(* Logix 5000 project; controller SmartManufacturingCell Emulate 5570 rev 33.11; software revision 33.03 *)
// Simulation only. Core cell candidate; acceptance pending.

TASK MainTask (periodic, rate 20 ms, priority 10, watchdog 500 ms) : Program_System, Program_Conveyor, Program_Filling, Program_Inspection, Program_Production, Program_Simulation

MODULES
   Local : Emulate 5570 (ICP 4, rev 33.11)
END_MODULES

TYPE UDT_Bottle :   // Bottle record
STRUCT
   Occupied : BOOL;   // A tracked bottle occupies this position
   FillComplete : BOOL;   // This bottle completed filling
   InspectionComplete : BOOL;   // This bottle has a valid inspection result
   RejectRequired : BOOL;   // Inspection determined this bottle must be rejected
END_STRUCT
END_TYPE

VAR_GLOBAL   (* controller tags *)
   Cfg_FillTimeMs : DINT := 1500;   // Fill duration; 100..3000 ms. Sampled when filling starts.
   Cfg_InspectionTimeMs : DINT := 500;   // Inspection duration; 100..2000 ms. Sampled when inspection starts.
   Conveyor_Flt_FailToStart : BOOL; {access Read Only}   // Conveyor commanded but running feedback missing for 2 s Latched; clear cell, remove cause, then fresh Reset.
   Conveyor_Sts_ResetAccepted : BOOL; {access Read Only}   // One-execution indication that conveyor fault reset was accepted.
   Exit_Flt_DischargeTimeout : BOOL; {access Read Only}   // Good or reject bottle departure not confirmed within 3 s Latched; clear cell, remove cause, then fresh Reset.
   Exit_Sts_GoodCompletePulse : BOOL; {access Read Only}   // Exit Sts GoodCompletePulse
   Exit_Sts_RejectCompletePulse : BOOL; {access Read Only}   // Exit Sts RejectCompletePulse
   Exit_Sts_ResetAccepted : BOOL; {access Read Only}   // Exit Sts ResetAccepted
   Exit_Sts_State : DINT; {access Read Only}   // 0 Empty; 10 Waiting; 20 Good discharge; 30 Extending; 40 Reject discharge; 50 Retracting; 60 Complete; 90 Faulted
   Filling_Flt_FillTimeout : BOOL; {access Read Only}   // Fill completion not received within 4 s Latched; clear cell, remove cause, then fresh Reset.
   Filling_Flt_ValveFailToClose : BOOL; {access Read Only}   // Fill valve did not close within 2 s Latched; clear cell, remove cause, then fresh Reset.
   Filling_Sts_ActiveFillTimeMs : DINT; {access Read Only}   // Sampled fill duration for current bottle
   Filling_Sts_ResetAccepted : BOOL; {access Read Only}   // Filling Sts ResetAccepted
   Filling_Sts_State : DINT; {access Read Only}   // 0 Empty; 10 Waiting; 20 Filling; 30 Closing; 40 Complete; 90 Faulted
   HMI_Cmd_Acknowledge : BOOL;   // Acknowledge alarm indication; does not reset faults
   HMI_Cmd_ClearCell : BOOL;   // Request removal of simulated bottles during fault recovery
   HMI_Cmd_ConveyorJog : BOOL;   // Request conveyor movement while held
   HMI_Cmd_FillValveOpen : BOOL;
   HMI_Cmd_LoadBottle : BOOL;   // Request one simulated bottle at the available entry position
   HMI_Cmd_RejectExtend : BOOL;
   HMI_Cmd_Reset : BOOL;   // Request fault reset after recovery conditions are satisfied
   HMI_Cmd_ResetStatistics : BOOL;   // Clear production statistics only when Stopped and cell empty
   HMI_Cmd_SelectAuto : BOOL;   // Request Auto mode
   HMI_Cmd_SelectManual : BOOL;   // Request Manual mode
   HMI_Cmd_Start : BOOL;   // Request automatic production start
   HMI_Cmd_Stop : BOOL;   // Request controlled production stop
   HMI_Sim_BottleMissingAtFill : BOOL;   // Suppress Fill photoeye while retaining simulated bottle presence. Simulation test only.
   HMI_Sim_ConveyorFailToStart : BOOL;   // Suppress conveyor running feedback. Simulation test only.
   HMI_Sim_FillFailToComplete : BOOL;   // Suppress simulated filling completion. Simulation test only.
   HMI_Sim_FillValveFailToClose : BOOL;   // Suppress fill valve closed feedback. Simulation test only.
   HMI_Sim_GoodDischargeJam : BOOL;   // Prevent good bottle departure. Simulation test only.
   HMI_Sim_IndexJam : BOOL;   // Prevent simulated index travel from completing. Simulation test only.
   HMI_Sim_IndexPositionMismatch : BOOL;   // Invert simulated Fill occupancy on transfer to test confirmation. Simulation test only.
   HMI_Sim_InspectionFailToComplete : BOOL;   // Prevent inspection process timer from completing. Simulation test only.
   HMI_Sim_NextInspectionRejects : BOOL;   // Select Reject for the next inspection
   HMI_Sim_RejectDischargeJam : BOOL;   // Prevent rejected bottle departure. Simulation test only.
   HMI_Sim_RejectFailToExtend : BOOL;   // Suppress reject extended feedback. Simulation test only.
   HMI_Sim_RejectFailToRetract : BOOL;   // Suppress reject retracted feedback. Simulation test only.
   Inspection_Flt_Timeout : BOOL; {access Read Only}   // Inspection did not finish within 3 s Latched; clear cell, remove cause, then fresh Reset.
   Inspection_Sts_ResetAccepted : BOOL; {access Read Only}   // Inspection Sts ResetAccepted
   Inspection_Sts_State : DINT; {access Read Only}   // 0 Empty; 10 Waiting; 20 Inspecting; 40 Complete; 90 Faulted
   Production_Bottles : UDT_Bottle[4]; {access Read Only}
   Production_Flt_IndexConfirmTimeout : BOOL; {access Read Only}   // Post-index positions not confirmed within 1 s Latched; clear cell, remove cause, then fresh Reset.
   Production_Flt_IndexInterlock : BOOL; {access Read Only}   // Movement interlock lost during indexing Latched; clear cell, remove cause, then fresh Reset.
   Production_Flt_IndexTimeout : BOOL; {access Read Only}   // Index completion not received within 3 s Latched; clear cell, remove cause, then fresh Reset.
   Production_Flt_InvalidConfiguration : BOOL; {access Read Only}   // Fill or inspection time outside permitted limits Latched; clear cell, remove cause, then fresh Reset.
   Production_Flt_InvalidState : BOOL; {access Read Only}   // Machine, sequence, station state, or mode combination invalid Latched; clear cell, remove cause, then fresh Reset.
   Production_Flt_StartupRecoveryRequired : BOOL; {access Read Only}   // Restart found bottles or interrupted activity Latched; clear cell, remove cause, then fresh Reset.
   Production_Flt_TrackingMismatch : BOOL; {access Read Only}   // Stationary bottle tracking and sensors disagree or processing history invalid Latched; clear cell, remove cause, then fresh Reset.
   Production_Stats_FaultSeconds : REAL; {access Read Only}   // FaultSeconds based on 20 ms scheduled executions; not a wall-clock historian.
   Production_Stats_GoodCount : DINT; {access Read Only}   // Retained GoodCount; count only confirmed departures (recovery losses separate).
   Production_Stats_LastCycleSeconds : REAL; {access Read Only}   // LastCycleSeconds based on 20 ms scheduled executions; not a wall-clock historian.
   Production_Stats_RatePerMinute : REAL; {access Read Only}   // RatePerMinute based on 20 ms scheduled executions; not a wall-clock historian.
   Production_Stats_RecoveryLossCount : DINT; {access Read Only}   // Retained RecoveryLossCount; count only confirmed departures (recovery losses separate).
   Production_Stats_RejectCount : DINT; {access Read Only}   // Retained RejectCount; count only confirmed departures (recovery losses separate).
   Production_Stats_RunSeconds : REAL; {access Read Only}   // RunSeconds based on 20 ms scheduled executions; not a wall-clock historian.
   Production_Stats_StoppedSeconds : REAL; {access Read Only}   // StoppedSeconds based on 20 ms scheduled executions; not a wall-clock historian.
   Production_Stats_TotalCount : DINT; {access Read Only}   // Retained TotalCount; count only confirmed departures (recovery losses separate).
   Production_Sts_ClearCellAccepted : BOOL; {access Read Only}
   Production_Sts_ClearCellAllowed : BOOL; {access Read Only}
   Production_Sts_CounterSaturated : BOOL; {access Read Only}   // Production Sts CounterSaturated
   Production_Sts_IndexAllowed : BOOL; {access Read Only}
   Production_Sts_IndexCommitted : BOOL; {access Read Only}   // Bottle records transferred for the current confirmed index; cleared outside ConfirmPositions.
   Production_Sts_IndexDemand : BOOL; {access Read Only}
   Production_Sts_IndexPositionsMatch : BOOL; {access Read Only}   // Post-index positions verified in ConfirmPositions with conveyor stopped.
   Production_Sts_LoadAccepted : BOOL; {access Read Only}
   Production_Sts_LoadAllowed : BOOL; {access Read Only}
   Production_Sts_LoadBlockReason : DINT; {access Read Only}   // 0 allowed; 10 not Auto Running/ProcessStations; 20 command conflict; 30 conveyor moving; 40 Entry occupied; 50 fault/startup incomplete
   Production_Sts_ResetAccepted : BOOL; {access Read Only}
   Production_Sts_SequenceState : DINT; {access Read Only}   // 0 = Idle 10 = ProcessStations 20 = Indexing 30 = ConfirmPositions
   Production_Sts_StationsReady : BOOL; {access Read Only}
   Reject_Flt_FailToExtend : BOOL;   // Reject actuator did not extend within 2 s Latched; clear cell, remove cause, then fresh Reset.
   Reject_Flt_FailToRetract : BOOL;   // Reject actuator did not retract within 2 s Latched; clear cell, remove cause, then fresh Reset.
   Reject_Sts_BlockReason : DINT; {access Read Only}   // Reason manual reject extension is unavailable. 0 = Ready to accept Extend. 10 = Release Extend to rearm. 20 = Good-bottle discharge active. 30 = Conveyor commanded or running. 40 = Stop request held. 50 = Machine is not Stopped. 60 = Mannual mode inactive or Auto Active. 70 = Blocking fault active. 99 = Permission unavailable for another reason.
   Reject_Sts_ResetAccepted : BOOL; {access Read Only}
   Sim_In_ConveyorRunning : BOOL; {access Read Only}   // Simulated conveyor movement feedback
   Sim_In_EntryPE : BOOL; {access Read Only}   // Simulated bottle detected at entry
   Sim_In_ExitPE : BOOL; {access Read Only}   // Simulated bottle detected at Reject/Exit position
   Sim_In_FillComplete : BOOL; {access Read Only}   // Sim In FillComplete
   Sim_In_FillPE : BOOL; {access Read Only}   // Simulated bottle detected at filling position
   Sim_In_FillValveClosed : BOOL; {access Read Only}   // Simulated fill valve confirmed closed
   Sim_In_GoodExitPE : BOOL; {access Read Only}   // Bottle detected passing through good discharge path
   Sim_In_IndexComplete : BOOL; {access Read Only}   // Simulated conveyor completed one station-spacing movement
   Sim_In_InspectionPE : BOOL; {access Read Only}   // Simulated bottle detected at inspection position
   Sim_In_RejectExitPE : BOOL; {access Read Only}   // Bottle detected passing through reject discharge path
   Sim_In_RejectExtended : BOOL; {access Read Only}   // Simulated reject actuator confirmed extended
   Sim_In_RejectRetracted : BOOL; {access Read Only}   // Simulated reject actuator confirmed retracted
   Sim_Out_ConveyorRun : BOOL; {access Read Only}   // Command simulated conveyor to run
   Sim_Out_FillValveOpen : BOOL; {access Read Only}   // Command simulated fill valve to open
   Sim_Out_GoodDischargeRun : BOOL; {access Read Only}   // Command simulated good-bottle discharge mechanism to run
   Sim_Out_RejectExtend : BOOL; {access Read Only}   // Command simulated reject actuator to extend
   Sim_Sts_BottlesPresent : BOOL; {access Read Only}   // Sim Sts BottlesPresent
   Sys_Sts_ActiveAlarmCount : DINT; {access Read Only}   // Number of active latched faults
   Sys_Sts_AlarmUnacknowledged : BOOL; {access Read Only}   // Sys Sts AlarmUnacknowledged
   Sys_Sts_AutoMode : BOOL; {access Read Only}   // Auto mode accepted and active
   Sys_Sts_BlockingFault : BOOL; {access Read Only}   // Active blocking fault prevents production and manual equipment operation.
   Sys_Sts_CellEmpty : BOOL; {access Read Only}   // Sys Sts CellEmpty
   Sys_Sts_EquipmentHome : BOOL; {access Read Only}   // Sys Sts EquipmentHome
   Sys_Sts_FirstFaultCode : DINT; {access Read Only}   // Lowest active fault code; zero means none
   Sys_Sts_InjectionsClear : BOOL; {access Read Only}   // Sys Sts InjectionsClear
   Sys_Sts_MachineState : DINT; {access Read Only}   // 0 = Stopped 10 = Running 20 = Stopping 30 = Faulted
   Sys_Sts_ManualMode : BOOL; {access Read Only}   // Manual mode accepted and active
   Sys_Sts_OperationsIdle : BOOL; {access Read Only}   // Sys Sts OperationsIdle
   Sys_Sts_ResetAllowed : BOOL; {access Read Only}   // Sys Sts ResetAllowed
   Sys_Sts_StartAllowed : BOOL; {access Read Only}
   Sys_Sts_StartupReady : BOOL; {access Read Only}   // Sys Sts StartupReady
END_VAR

PROGRAM Program_Conveyor   (* main routine MainRoutine *)
// Conveyor commands, movement permissives, and index monitoring.
VAR
   Conveyor_AutoRunAllowed : BOOL; {access None}
   Conveyor_JogArmed : BOOL; {access Read Only}
   Conveyor_ManualJogAllowed : BOOL; {access Read Only}   // Manual conveyor jog is permitted
   Conveyor_MovementAllowed : BOOL; {access Read Only}   // Equipment conditions permit conveyor movement
   ConveyorResetONS : BOOL; {access None}
   ConveyorStartTimeout : TIMER := (PRE := 2000);   // Non-retentive timer; preset in milliseconds.
END_VAR

ROUTINE Conveyor_Control   (* ladder *)
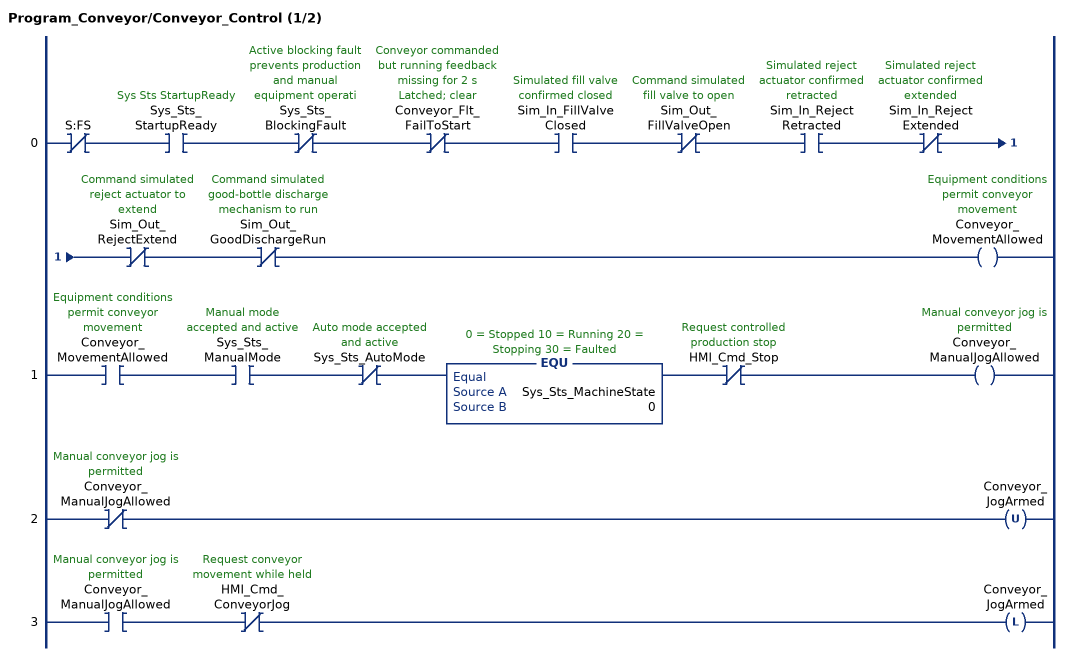
   0: XIO(S:FS)XIC(Sys_Sts_StartupReady)XIO(Sys_Sts_BlockingFault)XIO(Conveyor_Flt_FailToStart)XIC(Sim_In_FillValveClosed)XIO(Sim_Out_FillValveOpen)XIC(Sim_In_RejectRetracted)XIO(Sim_In_RejectExtended)XIO(Sim_Out_RejectExtend)XIO(Sim_Out_GoodDischargeRun)OTE(Conveyor_MovementAllowed);
   1: XIC(Conveyor_MovementAllowed)XIC(Sys_Sts_ManualMode)XIO(Sys_Sts_AutoMode)EQU(Sys_Sts_MachineState,0)XIO(HMI_Cmd_Stop)OTE(Conveyor_ManualJogAllowed);
   2: XIO(Conveyor_ManualJogAllowed)OTU(Conveyor_JogArmed);
   3: XIC(Conveyor_ManualJogAllowed)XIO(HMI_Cmd_ConveyorJog)OTL(Conveyor_JogArmed);
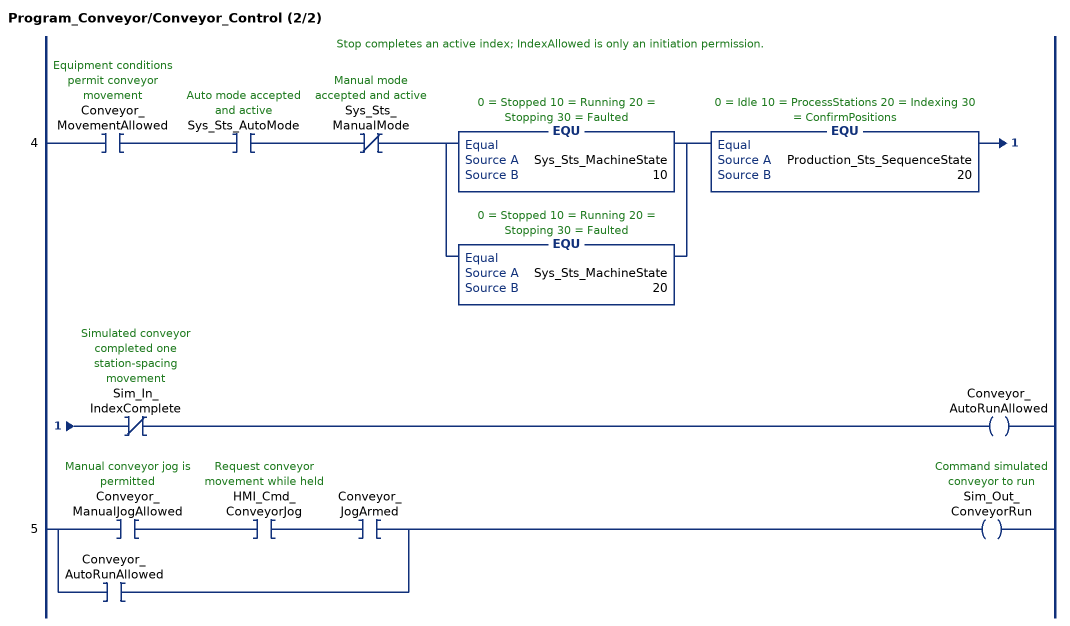
   // Stop completes an active index; IndexAllowed is only an initiation permission.
   4: XIC(Conveyor_MovementAllowed)XIC(Sys_Sts_AutoMode)XIO(Sys_Sts_ManualMode)[EQU(Sys_Sts_MachineState,10) ,EQU(Sys_Sts_MachineState,20) ]EQU(Production_Sts_SequenceState,20)XIO(Sim_In_IndexComplete)OTE(Conveyor_AutoRunAllowed);
   5: [XIC(Conveyor_ManualJogAllowed) XIC(HMI_Cmd_ConveyorJog) XIC(Conveyor_JogArmed) ,XIC(Conveyor_AutoRunAllowed) ]OTE(Sim_Out_ConveyorRun);
END_ROUTINE

ROUTINE Conveyor_Faults   (* ladder *)
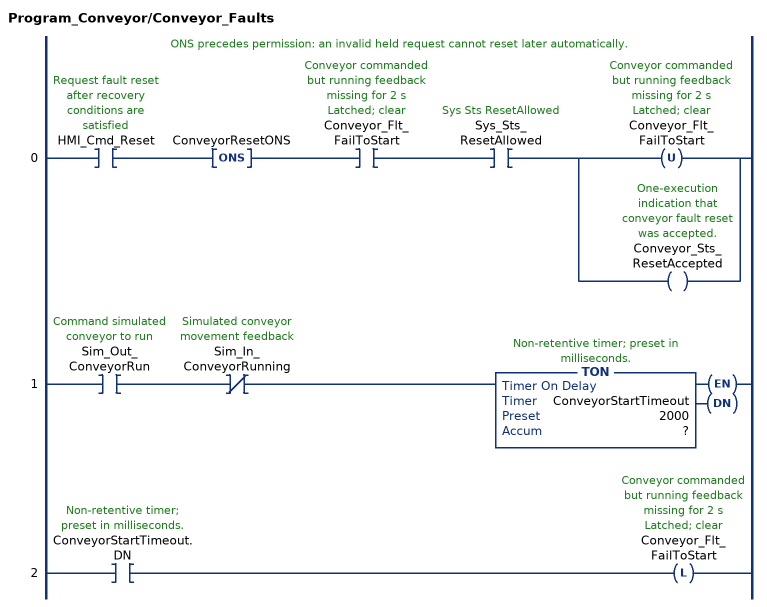
   // ONS precedes permission: an invalid held request cannot reset later automatically.
   0: XIC(HMI_Cmd_Reset)ONS(ConveyorResetONS)XIC(Conveyor_Flt_FailToStart)XIC(Sys_Sts_ResetAllowed)[OTU(Conveyor_Flt_FailToStart) ,OTE(Conveyor_Sts_ResetAccepted) ];
   1: XIC(Sim_Out_ConveyorRun)XIO(Sim_In_ConveyorRunning)TON(ConveyorStartTimeout,?,?);
   2: XIC(ConveyorStartTimeout.DN)OTL(Conveyor_Flt_FailToStart);
END_ROUTINE

ROUTINE MainRoutine   (* ladder *)
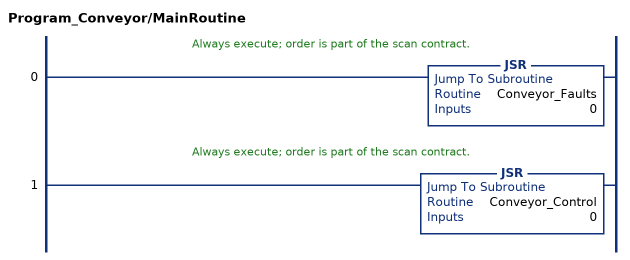
   // Always execute; order is part of the scan contract.
   0: JSR(Conveyor_Faults,0);
   // Always execute; order is part of the scan contract.
   1: JSR(Conveyor_Control,0);
END_ROUTINE
END_PROGRAM

PROGRAM Program_Filling   (* main routine MainRoutine *)
// Filling station valve control, timing, permissives, and faults.
VAR
   Fill_AutoOpenAllowed : BOOL; {access None}
   Fill_ManualOpenAllowed : BOOL; {access Read Only}
   Fill_ManualOpenArmed : BOOL; {access Read Only}
   Fill_StateAtScan : DINT; {access None}
   FillingResetONS : BOOL; {access None}
   FillProcessTimeout : TIMER := (PRE := 4000); {access None}   // Non-retentive timer; preset in milliseconds.
   FillValveCloseTimeout : TIMER := (PRE := 2000); {access None}   // Non-retentive timer; preset in milliseconds.
END_VAR

ROUTINE Filling_Control   (* ladder *)
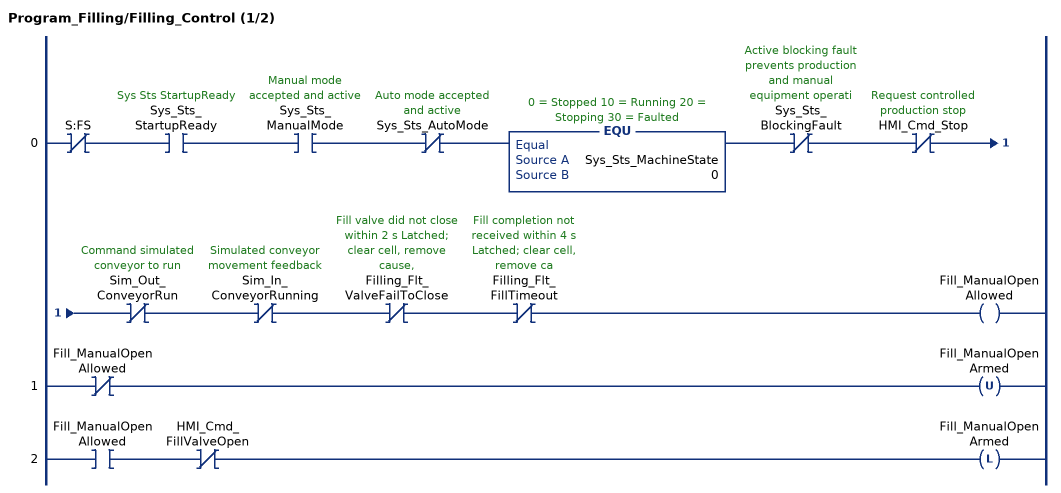
   0: XIO(S:FS)XIC(Sys_Sts_StartupReady)XIC(Sys_Sts_ManualMode)XIO(Sys_Sts_AutoMode)EQU(Sys_Sts_MachineState,0)XIO(Sys_Sts_BlockingFault)XIO(HMI_Cmd_Stop)XIO(Sim_Out_ConveyorRun)XIO(Sim_In_ConveyorRunning)XIO(Filling_Flt_ValveFailToClose)XIO(Filling_Flt_FillTimeout)OTE(Fill_ManualOpenAllowed);
   1: XIO(Fill_ManualOpenAllowed)OTU(Fill_ManualOpenArmed);
   2: XIC(Fill_ManualOpenAllowed)XIO(HMI_Cmd_FillValveOpen)OTL(Fill_ManualOpenArmed);
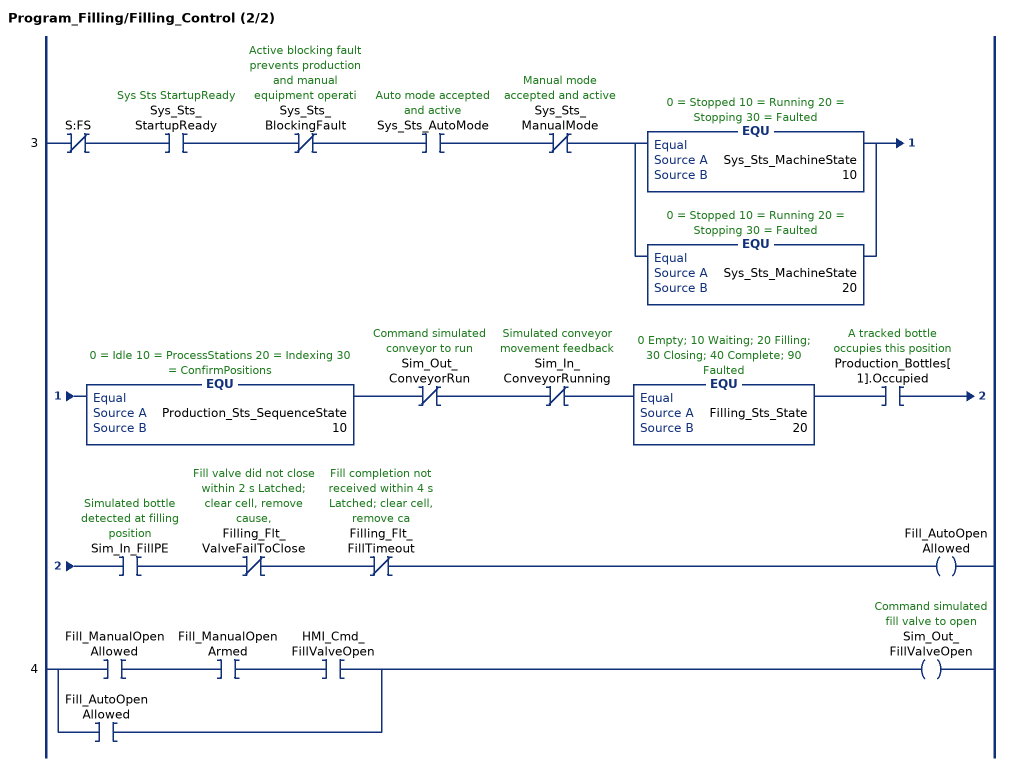
   3: XIO(S:FS)XIC(Sys_Sts_StartupReady)XIO(Sys_Sts_BlockingFault)XIC(Sys_Sts_AutoMode)XIO(Sys_Sts_ManualMode)[EQU(Sys_Sts_MachineState,10) ,EQU(Sys_Sts_MachineState,20) ]EQU(Production_Sts_SequenceState,10)XIO(Sim_Out_ConveyorRun)XIO(Sim_In_ConveyorRunning)EQU(Filling_Sts_State,20)XIC(Production_Bottles[1].Occupied)XIC(Sim_In_FillPE)XIO(Filling_Flt_ValveFailToClose)XIO(Filling_Flt_FillTimeout)OTE(Fill_AutoOpenAllowed);
   4: [XIC(Fill_ManualOpenAllowed) XIC(Fill_ManualOpenArmed) XIC(HMI_Cmd_FillValveOpen) ,XIC(Fill_AutoOpenAllowed) ]OTE(Sim_Out_FillValveOpen);
END_ROUTINE

ROUTINE Filling_Faults   (* ladder *)
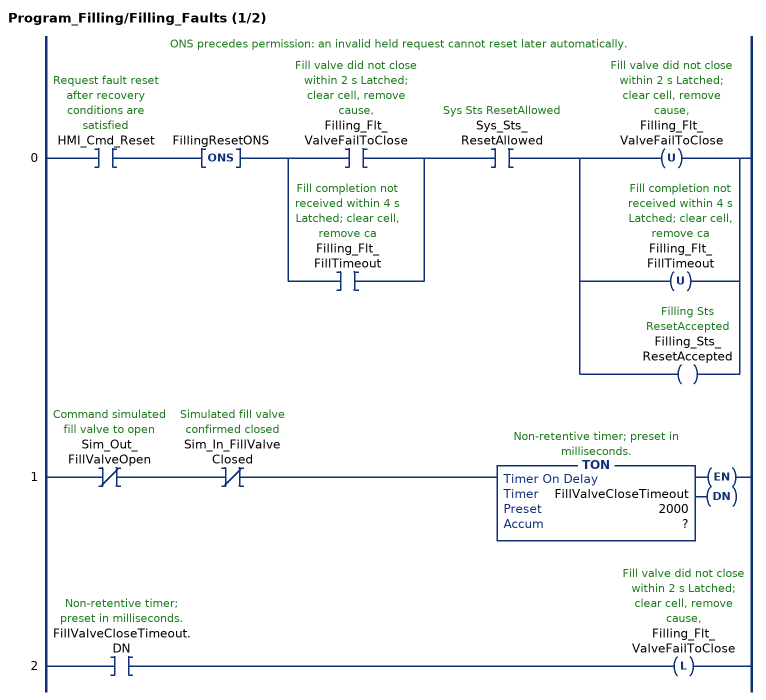
   // ONS precedes permission: an invalid held request cannot reset later automatically.
   0: XIC(HMI_Cmd_Reset)ONS(FillingResetONS)[XIC(Filling_Flt_ValveFailToClose) ,XIC(Filling_Flt_FillTimeout) ]XIC(Sys_Sts_ResetAllowed)[OTU(Filling_Flt_ValveFailToClose) ,OTU(Filling_Flt_FillTimeout) ,OTE(Filling_Sts_ResetAccepted) ];
   1: XIO(Sim_Out_FillValveOpen)XIO(Sim_In_FillValveClosed)TON(FillValveCloseTimeout,?,?);
   2: XIC(FillValveCloseTimeout.DN)OTL(Filling_Flt_ValveFailToClose);
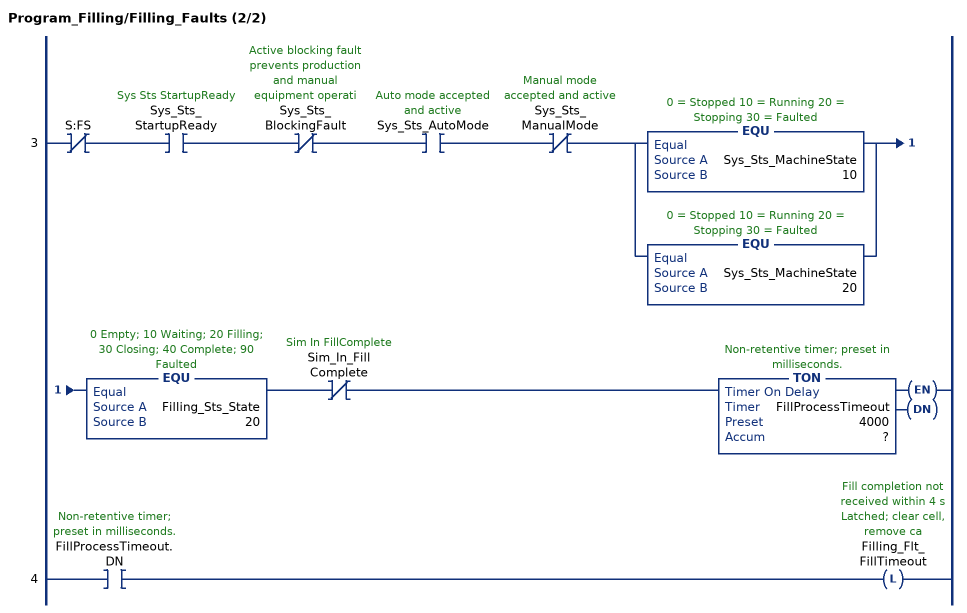
   3: XIO(S:FS)XIC(Sys_Sts_StartupReady)XIO(Sys_Sts_BlockingFault)XIC(Sys_Sts_AutoMode)XIO(Sys_Sts_ManualMode)[EQU(Sys_Sts_MachineState,10) ,EQU(Sys_Sts_MachineState,20) ]EQU(Filling_Sts_State,20)XIO(Sim_In_FillComplete)TON(FillProcessTimeout,?,?);
   4: XIC(FillProcessTimeout.DN)OTL(Filling_Flt_FillTimeout);
END_ROUTINE

ROUTINE Filling_Sequence   (* ladder *)
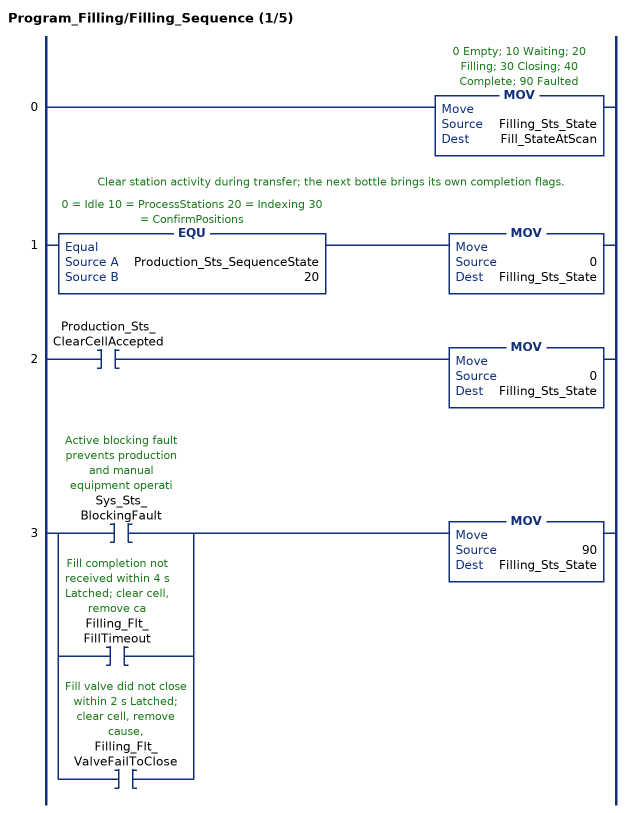
   0: MOV(Filling_Sts_State,Fill_StateAtScan);
   // Clear station activity during transfer; the next bottle brings its own completion flags.
   1: EQU(Production_Sts_SequenceState,20)MOV(0,Filling_Sts_State);
   2: XIC(Production_Sts_ClearCellAccepted)MOV(0,Filling_Sts_State);
   3: [XIC(Sys_Sts_BlockingFault) ,XIC(Filling_Flt_FillTimeout) ,XIC(Filling_Flt_ValveFailToClose) ]MOV(90,Filling_Sts_State);
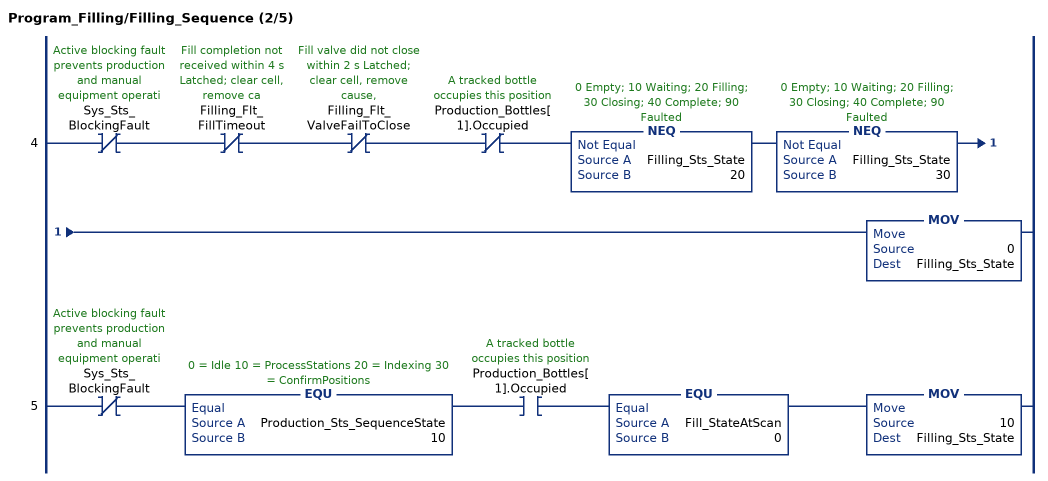
   4: XIO(Sys_Sts_BlockingFault)XIO(Filling_Flt_FillTimeout)XIO(Filling_Flt_ValveFailToClose)XIO(Production_Bottles[1].Occupied)NEQ(Filling_Sts_State,20)NEQ(Filling_Sts_State,30)MOV(0,Filling_Sts_State);
   5: XIO(Sys_Sts_BlockingFault)EQU(Production_Sts_SequenceState,10)XIC(Production_Bottles[1].Occupied)EQU(Fill_StateAtScan,0)MOV(10,Filling_Sts_State);
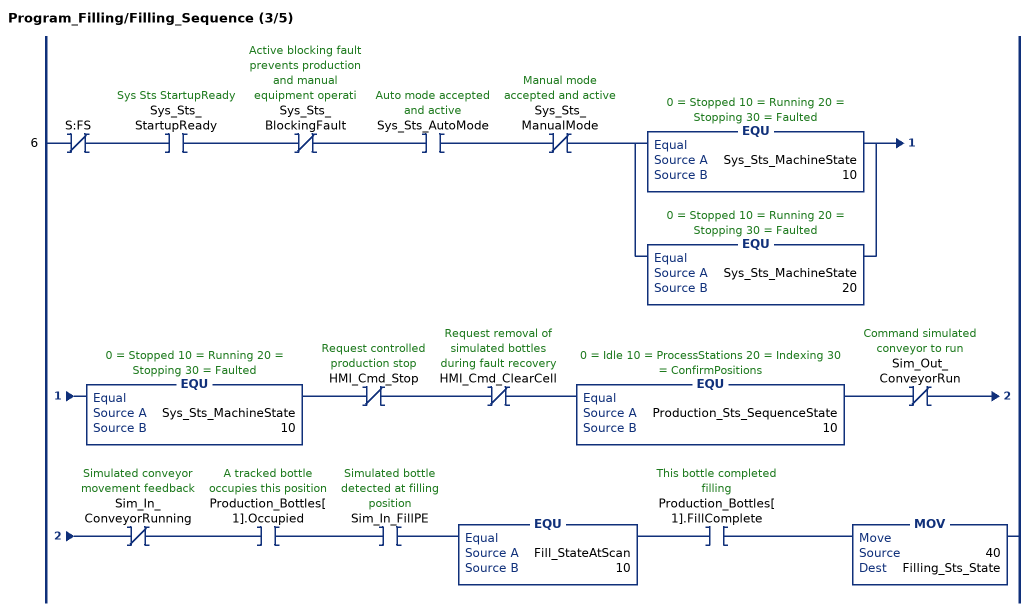
   6: XIO(S:FS)XIC(Sys_Sts_StartupReady)XIO(Sys_Sts_BlockingFault)XIC(Sys_Sts_AutoMode)XIO(Sys_Sts_ManualMode)[EQU(Sys_Sts_MachineState,10) ,EQU(Sys_Sts_MachineState,20) ]EQU(Sys_Sts_MachineState,10)XIO(HMI_Cmd_Stop)XIO(HMI_Cmd_ClearCell)EQU(Production_Sts_SequenceState,10)XIO(Sim_Out_ConveyorRun)XIO(Sim_In_ConveyorRunning)XIC(Production_Bottles[1].Occupied)XIC(Sim_In_FillPE)EQU(Fill_StateAtScan,10)XIC(Production_Bottles[1].FillComplete)MOV(40,Filling_Sts_State);
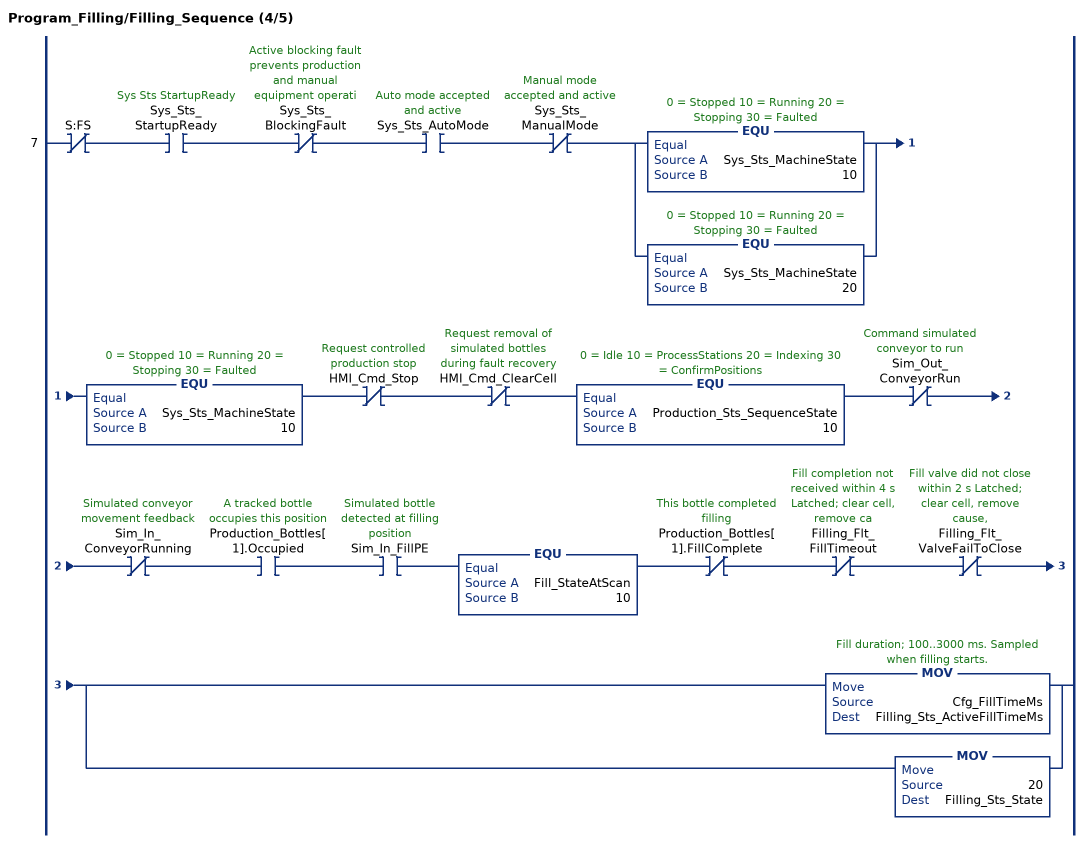
   7: XIO(S:FS)XIC(Sys_Sts_StartupReady)XIO(Sys_Sts_BlockingFault)XIC(Sys_Sts_AutoMode)XIO(Sys_Sts_ManualMode)[EQU(Sys_Sts_MachineState,10) ,EQU(Sys_Sts_MachineState,20) ]EQU(Sys_Sts_MachineState,10)XIO(HMI_Cmd_Stop)XIO(HMI_Cmd_ClearCell)EQU(Production_Sts_SequenceState,10)XIO(Sim_Out_ConveyorRun)XIO(Sim_In_ConveyorRunning)XIC(Production_Bottles[1].Occupied)XIC(Sim_In_FillPE)EQU(Fill_StateAtScan,10)XIO(Production_Bottles[1].FillComplete)XIO(Filling_Flt_FillTimeout)XIO(Filling_Flt_ValveFailToClose)[MOV(Cfg_FillTimeMs,Filling_Sts_ActiveFillTimeMs) ,MOV(20,Filling_Sts_State) ];
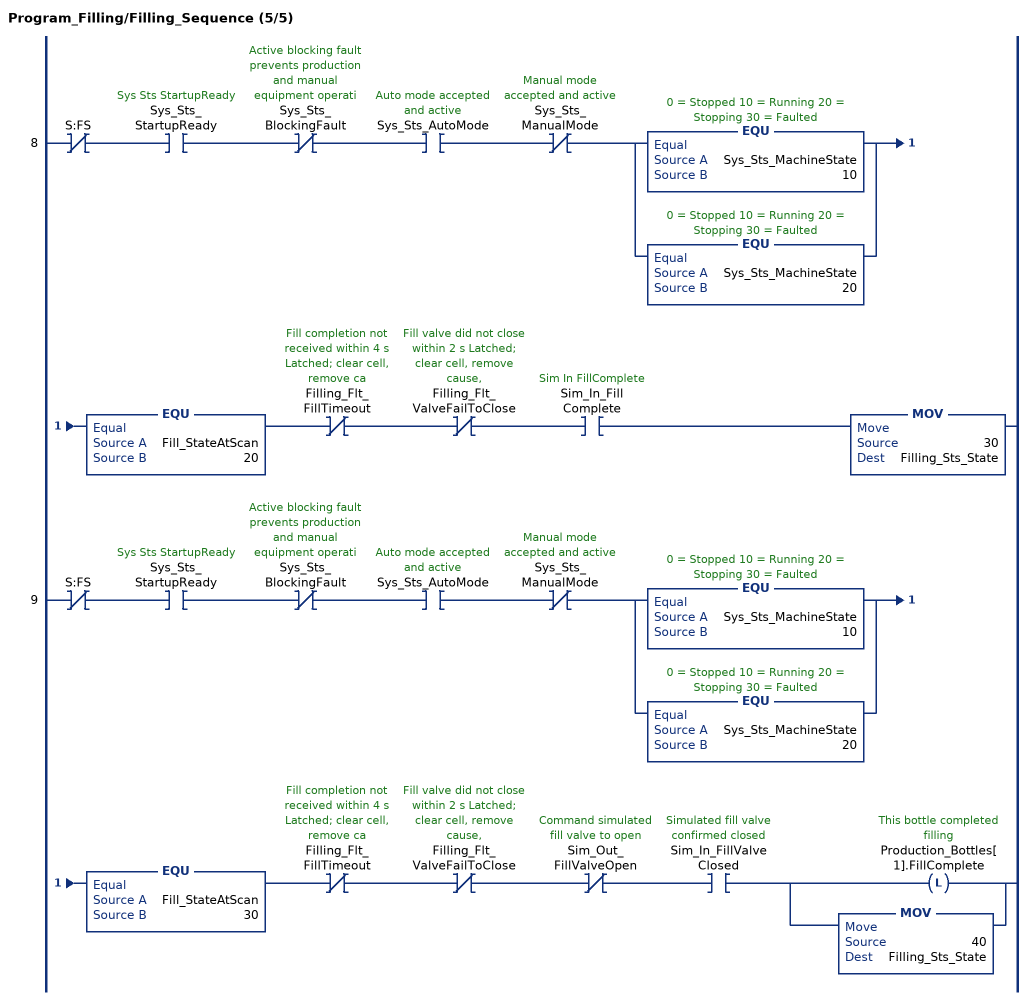
   8: XIO(S:FS)XIC(Sys_Sts_StartupReady)XIO(Sys_Sts_BlockingFault)XIC(Sys_Sts_AutoMode)XIO(Sys_Sts_ManualMode)[EQU(Sys_Sts_MachineState,10) ,EQU(Sys_Sts_MachineState,20) ]EQU(Fill_StateAtScan,20)XIO(Filling_Flt_FillTimeout)XIO(Filling_Flt_ValveFailToClose)XIC(Sim_In_FillComplete)MOV(30,Filling_Sts_State);
   9: XIO(S:FS)XIC(Sys_Sts_StartupReady)XIO(Sys_Sts_BlockingFault)XIC(Sys_Sts_AutoMode)XIO(Sys_Sts_ManualMode)[EQU(Sys_Sts_MachineState,10) ,EQU(Sys_Sts_MachineState,20) ]EQU(Fill_StateAtScan,30)XIO(Filling_Flt_FillTimeout)XIO(Filling_Flt_ValveFailToClose)XIO(Sim_Out_FillValveOpen)XIC(Sim_In_FillValveClosed)[OTL(Production_Bottles[1].FillComplete) ,MOV(40,Filling_Sts_State) ];
END_ROUTINE

ROUTINE MainRoutine   (* ladder *)
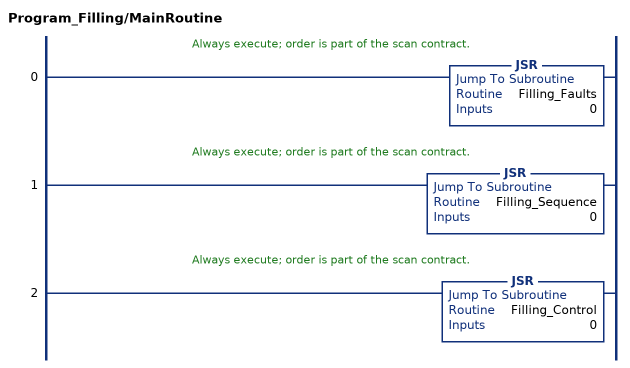
   // Always execute; order is part of the scan contract.
   0: JSR(Filling_Faults,0);
   // Always execute; order is part of the scan contract.
   1: JSR(Filling_Sequence,0);
   // Always execute; order is part of the scan contract.
   2: JSR(Filling_Control,0);
END_ROUTINE
END_PROGRAM

PROGRAM Program_Inspection   (* main routine MainRoutine *)
// Simulated inspection, reject actuator, and bottle discharge control.
VAR
   Exit_StateAtScan : DINT; {access None}
   ExitDischargeTimeout : TIMER := (PRE := 3000); {access None}   // Non-retentive timer; preset in milliseconds.
   ExitResetONS : BOOL; {access None}
   Inspection_RejectSample : BOOL; {access None}
   Inspection_StateAtScan : DINT; {access None}
   InspectionProcessDelay : TIMER := (PRE := 500); {access None}   // Non-retentive timer; preset in milliseconds.
   InspectionResetONS : BOOL; {access None}
   InspectionTimeout : TIMER := (PRE := 3000); {access None}   // Non-retentive timer; preset in milliseconds.
   Reject_AutoExtendAllowed : BOOL; {access None}
   Reject_ManualExtendAllowed : BOOL; {access Read Only}
   Reject_ManualExtendArmed : BOOL; {access Read Only}
   Reject_ResetAllowed : BOOL; {access None}   // Reject recovery conditions satisfied; permits a fresh Reset request.
   RejectExtendTimeout : TIMER := (PRE := 2000); {access None}   // Non-retentive timer; preset in milliseconds.
   RejectResetONS : BOOL; {access None}
   RejectRetractTimeout : TIMER := (PRE := 2000); {access None}   // Non-retentive timer; preset in milliseconds.
END_VAR

ROUTINE Exit_Control   (* ladder *)
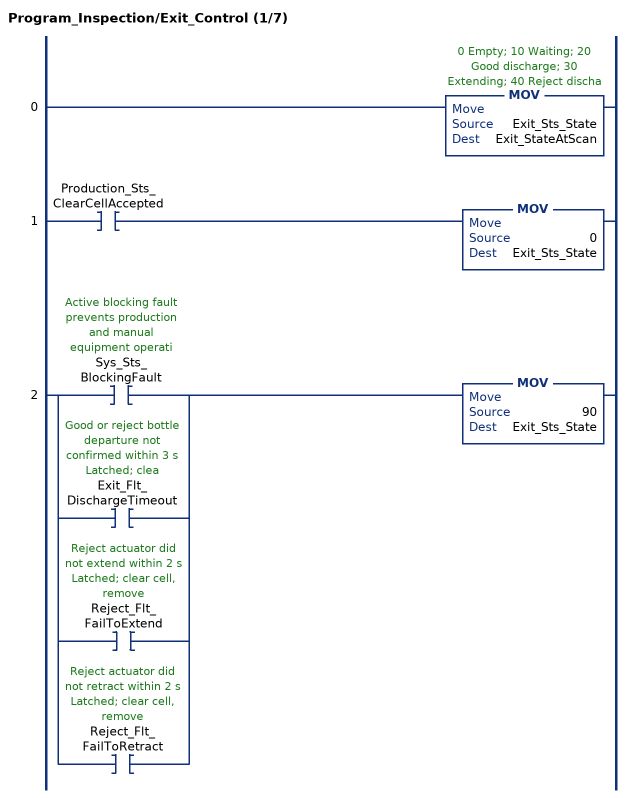
   0: MOV(Exit_Sts_State,Exit_StateAtScan);
   1: XIC(Production_Sts_ClearCellAccepted)MOV(0,Exit_Sts_State);
   2: [XIC(Sys_Sts_BlockingFault) ,XIC(Exit_Flt_DischargeTimeout) ,XIC(Reject_Flt_FailToExtend) ,XIC(Reject_Flt_FailToRetract) ]MOV(90,Exit_Sts_State);
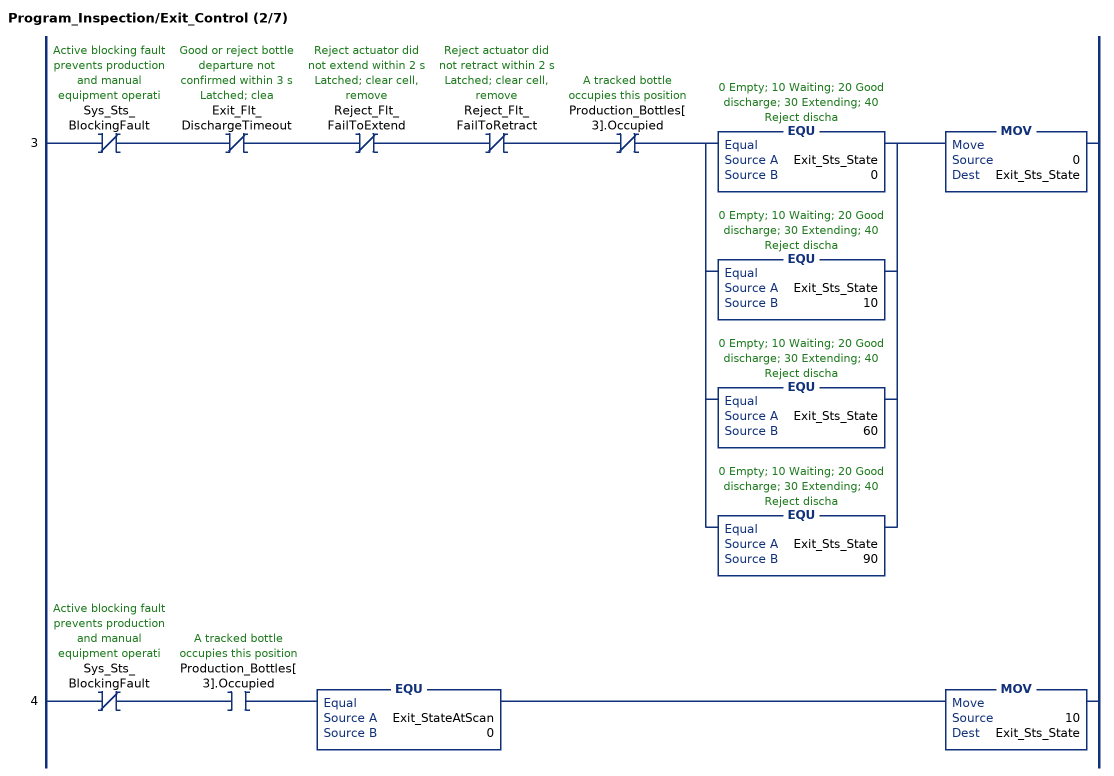
   3: XIO(Sys_Sts_BlockingFault)XIO(Exit_Flt_DischargeTimeout)XIO(Reject_Flt_FailToExtend)XIO(Reject_Flt_FailToRetract)XIO(Production_Bottles[3].Occupied)[EQU(Exit_Sts_State,0) ,EQU(Exit_Sts_State,10) ,EQU(Exit_Sts_State,60) ,EQU(Exit_Sts_State,90) ]MOV(0,Exit_Sts_State);
   4: XIO(Sys_Sts_BlockingFault)XIC(Production_Bottles[3].Occupied)EQU(Exit_StateAtScan,0)MOV(10,Exit_Sts_State);
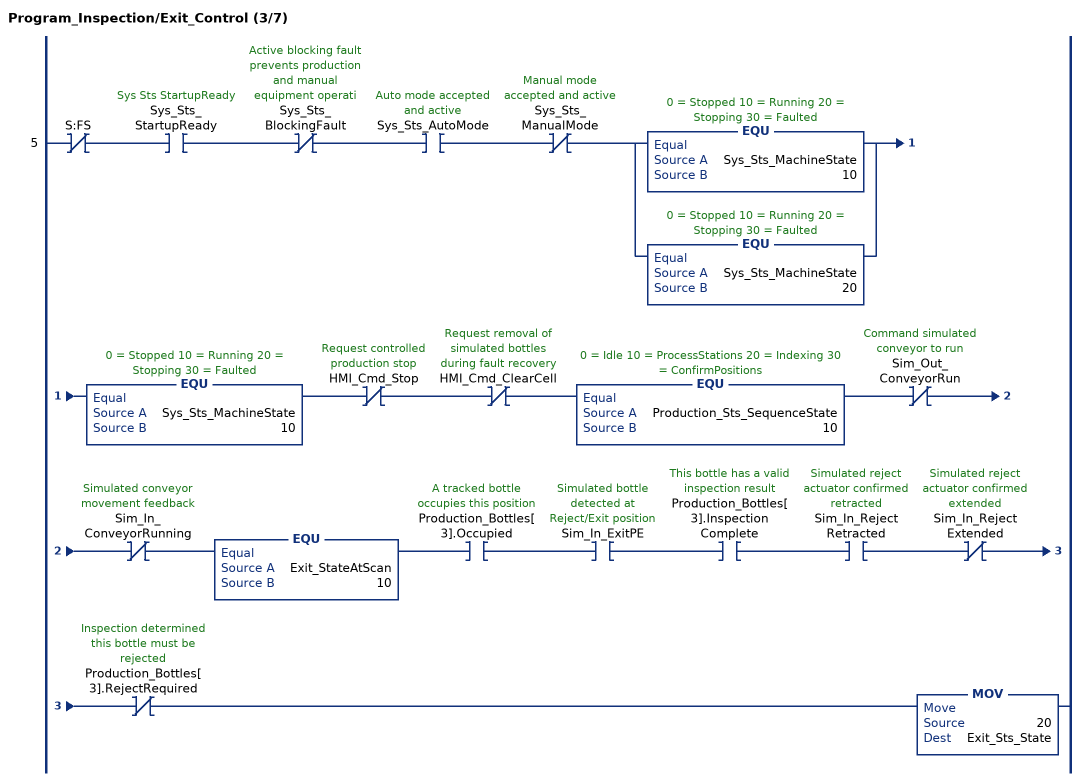
   5: XIO(S:FS)XIC(Sys_Sts_StartupReady)XIO(Sys_Sts_BlockingFault)XIC(Sys_Sts_AutoMode)XIO(Sys_Sts_ManualMode)[EQU(Sys_Sts_MachineState,10) ,EQU(Sys_Sts_MachineState,20) ]EQU(Sys_Sts_MachineState,10)XIO(HMI_Cmd_Stop)XIO(HMI_Cmd_ClearCell)EQU(Production_Sts_SequenceState,10)XIO(Sim_Out_ConveyorRun)XIO(Sim_In_ConveyorRunning)EQU(Exit_StateAtScan,10)XIC(Production_Bottles[3].Occupied)XIC(Sim_In_ExitPE)XIC(Production_Bottles[3].InspectionComplete)XIC(Sim_In_RejectRetracted)XIO(Sim_In_RejectExtended)XIO(Production_Bottles[3].RejectRequired)MOV(20,Exit_Sts_State);
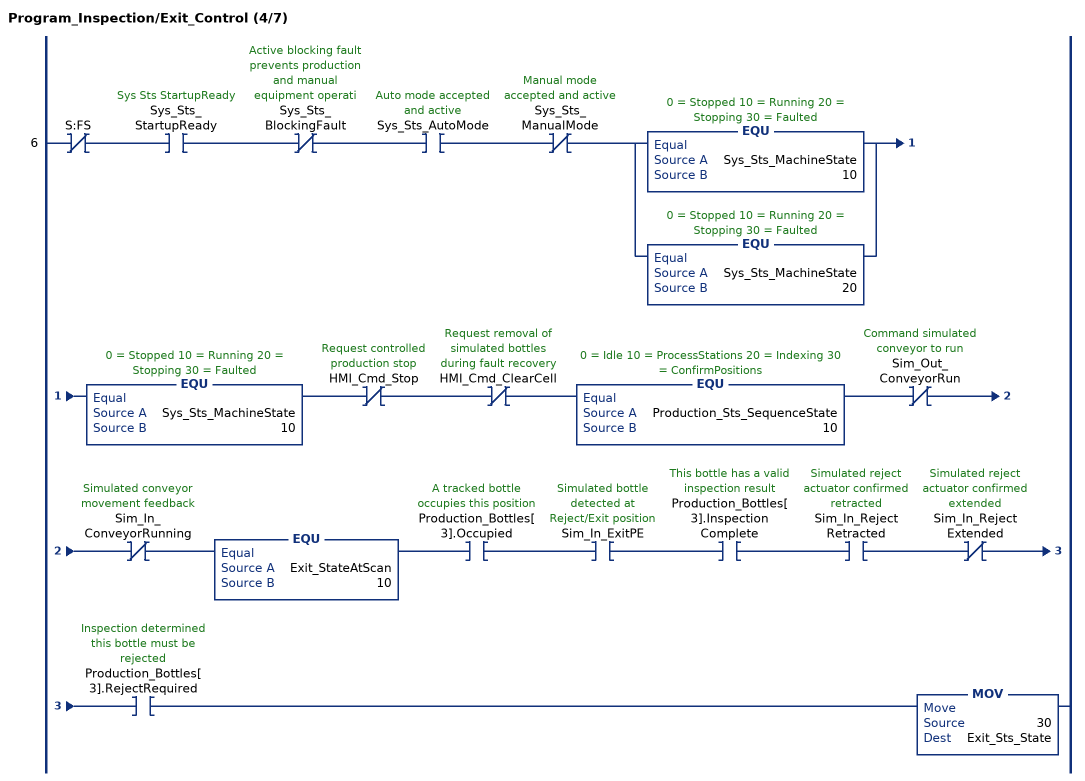
   6: XIO(S:FS)XIC(Sys_Sts_StartupReady)XIO(Sys_Sts_BlockingFault)XIC(Sys_Sts_AutoMode)XIO(Sys_Sts_ManualMode)[EQU(Sys_Sts_MachineState,10) ,EQU(Sys_Sts_MachineState,20) ]EQU(Sys_Sts_MachineState,10)XIO(HMI_Cmd_Stop)XIO(HMI_Cmd_ClearCell)EQU(Production_Sts_SequenceState,10)XIO(Sim_Out_ConveyorRun)XIO(Sim_In_ConveyorRunning)EQU(Exit_StateAtScan,10)XIC(Production_Bottles[3].Occupied)XIC(Sim_In_ExitPE)XIC(Production_Bottles[3].InspectionComplete)XIC(Sim_In_RejectRetracted)XIO(Sim_In_RejectExtended)XIC(Production_Bottles[3].RejectRequired)MOV(30,Exit_Sts_State);
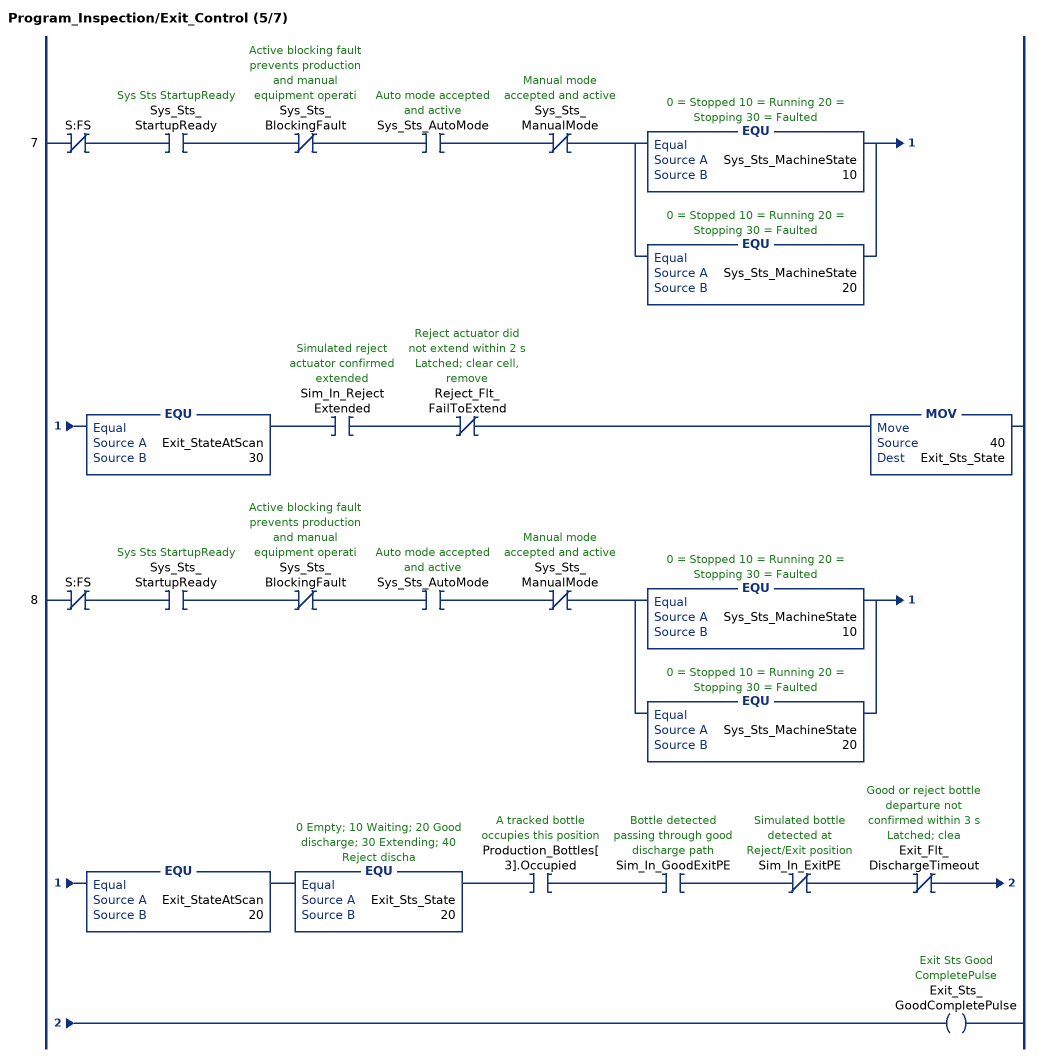
   7: XIO(S:FS)XIC(Sys_Sts_StartupReady)XIO(Sys_Sts_BlockingFault)XIC(Sys_Sts_AutoMode)XIO(Sys_Sts_ManualMode)[EQU(Sys_Sts_MachineState,10) ,EQU(Sys_Sts_MachineState,20) ]EQU(Exit_StateAtScan,30)XIC(Sim_In_RejectExtended)XIO(Reject_Flt_FailToExtend)MOV(40,Exit_Sts_State);
   8: XIO(S:FS)XIC(Sys_Sts_StartupReady)XIO(Sys_Sts_BlockingFault)XIC(Sys_Sts_AutoMode)XIO(Sys_Sts_ManualMode)[EQU(Sys_Sts_MachineState,10) ,EQU(Sys_Sts_MachineState,20) ]EQU(Exit_StateAtScan,20)EQU(Exit_Sts_State,20)XIC(Production_Bottles[3].Occupied)XIC(Sim_In_GoodExitPE)XIO(Sim_In_ExitPE)XIO(Exit_Flt_DischargeTimeout)OTE(Exit_Sts_GoodCompletePulse);
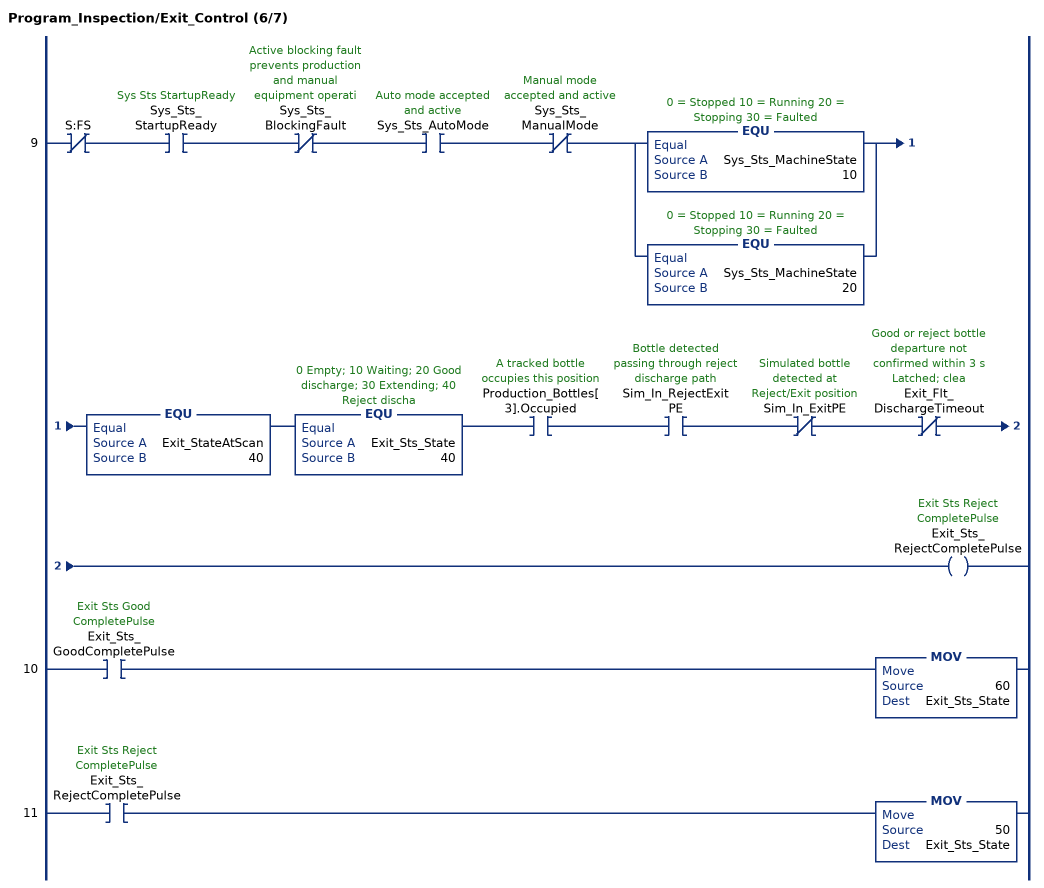
   9: XIO(S:FS)XIC(Sys_Sts_StartupReady)XIO(Sys_Sts_BlockingFault)XIC(Sys_Sts_AutoMode)XIO(Sys_Sts_ManualMode)[EQU(Sys_Sts_MachineState,10) ,EQU(Sys_Sts_MachineState,20) ]EQU(Exit_StateAtScan,40)EQU(Exit_Sts_State,40)XIC(Production_Bottles[3].Occupied)XIC(Sim_In_RejectExitPE)XIO(Sim_In_ExitPE)XIO(Exit_Flt_DischargeTimeout)OTE(Exit_Sts_RejectCompletePulse);
   10: XIC(Exit_Sts_GoodCompletePulse)MOV(60,Exit_Sts_State);
   11: XIC(Exit_Sts_RejectCompletePulse)MOV(50,Exit_Sts_State);
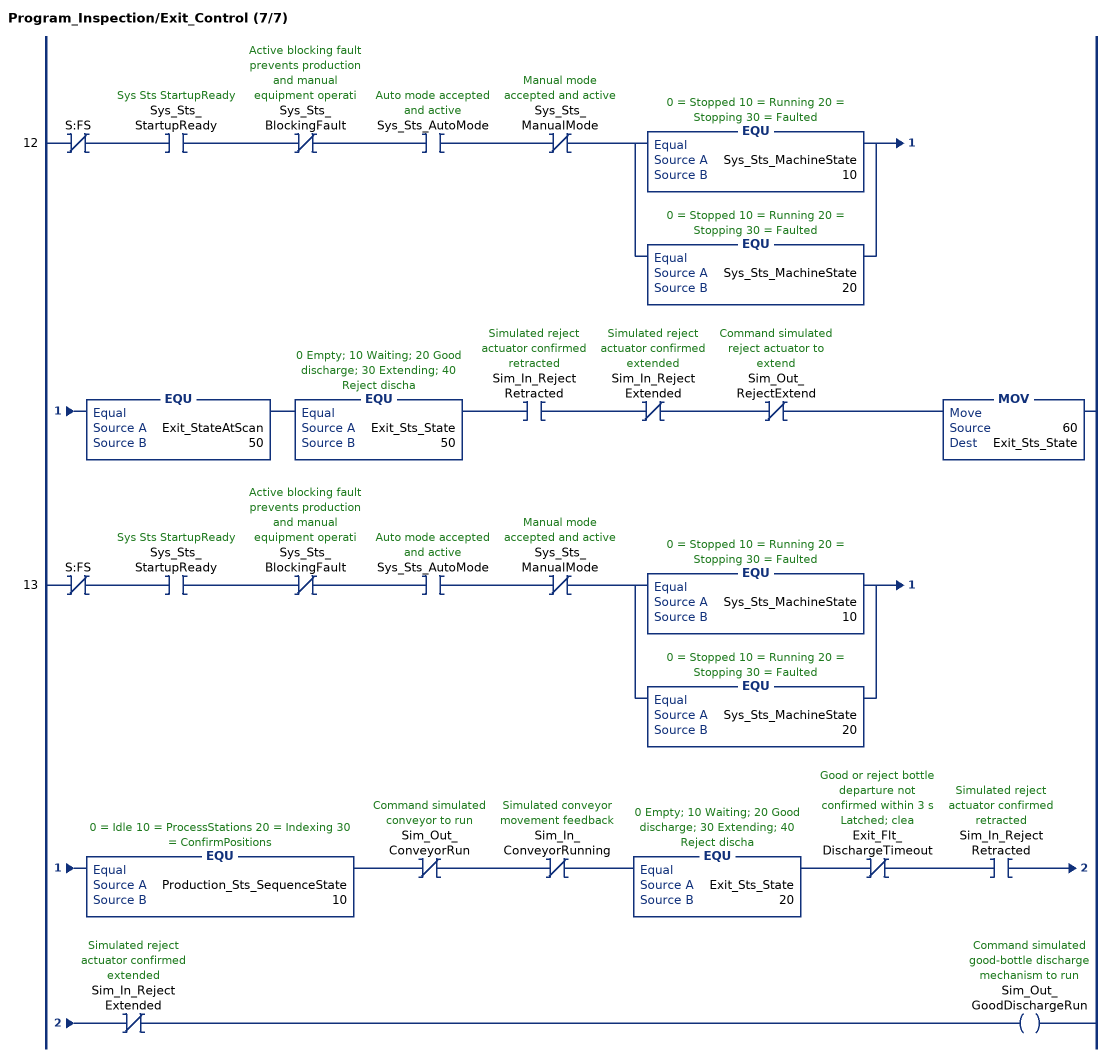
   12: XIO(S:FS)XIC(Sys_Sts_StartupReady)XIO(Sys_Sts_BlockingFault)XIC(Sys_Sts_AutoMode)XIO(Sys_Sts_ManualMode)[EQU(Sys_Sts_MachineState,10) ,EQU(Sys_Sts_MachineState,20) ]EQU(Exit_StateAtScan,50)EQU(Exit_Sts_State,50)XIC(Sim_In_RejectRetracted)XIO(Sim_In_RejectExtended)XIO(Sim_Out_RejectExtend)MOV(60,Exit_Sts_State);
   13: XIO(S:FS)XIC(Sys_Sts_StartupReady)XIO(Sys_Sts_BlockingFault)XIC(Sys_Sts_AutoMode)XIO(Sys_Sts_ManualMode)[EQU(Sys_Sts_MachineState,10) ,EQU(Sys_Sts_MachineState,20) ]EQU(Production_Sts_SequenceState,10)XIO(Sim_Out_ConveyorRun)XIO(Sim_In_ConveyorRunning)EQU(Exit_Sts_State,20)XIO(Exit_Flt_DischargeTimeout)XIC(Sim_In_RejectRetracted)XIO(Sim_In_RejectExtended)OTE(Sim_Out_GoodDischargeRun);
END_ROUTINE
